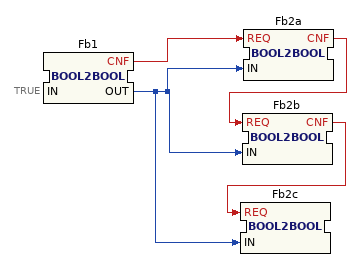
      [picture p24: application _03_DataConnections.Ex2b]
      FBS
        Fb1 : BOOL2BOOL(IN := TRUE);
        Fb2a : BOOL2BOOL;
        Fb2b : BOOL2BOOL;
        Fb2c : BOOL2BOOL;
      END_FBS
      EVENT_CONNECTIONS
        Fb1.CNF TO Fb2a.REQ;
        Fb2a.CNF TO Fb2b.REQ;
        Fb2b.CNF TO Fb2c.REQ;
      END_CONNECTIONS
      DATA_CONNECTIONS
        Fb1.OUT TO Fb2a.IN;
        Fb1.OUT TO Fb2b.IN;
        Fb1.OUT TO Fb2c.IN;
      END_CONNECTIONS
    END_SUBAPPLICATION
    SUBAPPLICATION Ex4b (* type casts (explicit, downcast) &#10;- trigger Fb1.REQ &#10;- expect Fb3.CUO and CV:=1 and Q:=TRUE *)
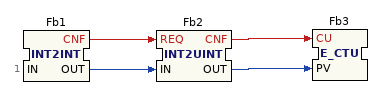
      FBS
        Fb1 : INT2INT(IN := 1);
        Fb3 : E_CTU;
        Fb2 : INT2UINT;
      END_FBS
      EVENT_CONNECTIONS
        Fb1.CNF TO Fb2.REQ;
        Fb2.CNF TO Fb3.CU;
      END_CONNECTIONS
      DATA_CONNECTIONS
        Fb1.OUT TO Fb2.IN;
        Fb2.OUT TO Fb3.PV;
      END_CONNECTIONS
    END_SUBAPPLICATION
    SUBAPPLICATION Ex5a (* type casts (implicit, upcast from UINT to LREAL) &#10;- trigger Fb1.CU  &#10;- expect Fb2.CNF and Fb2.OUT:=INT#6 *)
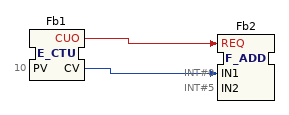
      FBS
        Fb1 : E_CTU(PV := 10);
        Fb2 : F_ADD(IN1 := INT#0, IN2 := INT#5);
      END_FBS
      EVENT_CONNECTIONS
        Fb1.CUO TO Fb2.REQ;
      END_CONNECTIONS
      DATA_CONNECTIONS
        Fb1.CV TO Fb2.IN1;
      END_CONNECTIONS
    END_SUBAPPLICATION
    SUBAPPLICATION Ex5b (* type casts (implicit, upcast from UINT to ANY_MAG) &#10;- trigger Fb1.CU &#10;- expect Fb2.CNF and Fb2.OUT:=REAL#1.0 *)
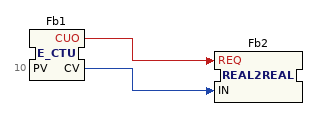
      FBS
        Fb1 : E_CTU(PV := 10);
        Fb2 : REAL2REAL;
      END_FBS
      EVENT_CONNECTIONS
        Fb1.CUO TO Fb2.REQ;
      END_CONNECTIONS
      DATA_CONNECTIONS
        Fb1.CV TO Fb2.IN;
      END_CONNECTIONS
    END_SUBAPPLICATION
  END_APPLICATION
  APPLICATION _07_Subapplications
    (* Group __Group01: connection to the interface *)
  END_APPLICATION
  APPLICATION _06_CompositeFBs
    (* Group __Group01: WITH bei composite FBs *)
  END_APPLICATION
  APPLICATION _02_Parameters
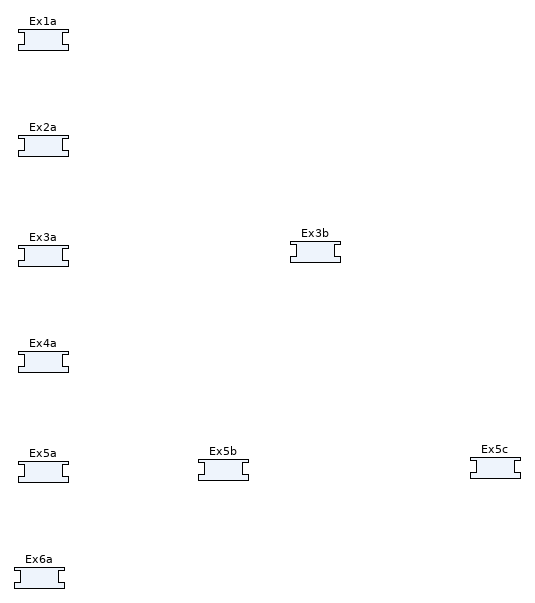
    (* Group Info_Parameters: The subapps in this App serve as test cases for various versions of parameters: &#10;- simple boolean parameters (including counter-examples) &#10;- initial value taken from type when no parameter is present &#10;- parameters with prefixes &#10;- upcasts in parameters *)
    SUBAPPLICATION Ex2a (* Parameters &#10; &#10;- Trigger EI  &#10;- Expect nothing *)
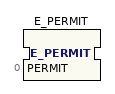
      FBS
        E_PERMIT : E_PERMIT(PERMIT := 0);
      END_FBS
    END_SUBAPPLICATION
    SUBAPPLICATION Ex1a (* Parameters overriding initial value of data type &#10; &#10;- Trigger E_PERMIT.EI  &#10;- Expect E_PERMIT.EO *)
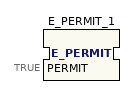
      FBS
        E_PERMIT_1 : E_PERMIT(PERMIT := TRUE);
      END_FBS
    END_SUBAPPLICATION
    SUBAPPLICATION Ex3a (* Initial Value (from type) &#10; &#10;- Trigger EI  &#10;- Expect EO *)
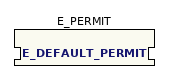
      FBS
        E_PERMIT : E_DEFAULT_PERMIT;
      END_FBS
    END_SUBAPPLICATION
    SUBAPPLICATION Ex4a (* Override initial value (from type) with parameter &#10; &#10;- Trigger EI  &#10;- Expect nothing *)
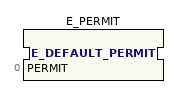
      FBS
        E_PERMIT : E_DEFAULT_PERMIT(PERMIT := 0);
      END_FBS
    END_SUBAPPLICATION
    SUBAPPLICATION Ex6a (* Any type: required casts  &#10; &#10;- Trigger REQ &#10;- Expect CNF and OUT:=13 *)
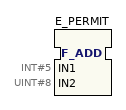
      FBS
        E_PERMIT : F_ADD(IN1 := INT#5, IN2 := UINT#8);
      END_FBS
    END_SUBAPPLICATION
    SUBAPPLICATION Ex5a (* integer parameter &#10; &#10;- Trigger REQ &#10;- Expect CNF, OUT:=5 *)
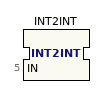
      FBS
        INT2INT : INT2INT(IN := 5);
      END_FBS
    END_SUBAPPLICATION
    SUBAPPLICATION Ex5b (* integer parameter with prefix &#10; &#10;- Trigger REQ &#10;- Expect CNF, OUT:=5 *)
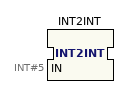
      FBS
        INT2INT : INT2INT(IN := INT#5);
      END_FBS
    END_SUBAPPLICATION
    SUBAPPLICATION Ex5c (* integer parameter with prefix (upcast) &#10; &#10;- Trigger REQ &#10;- Expect CNF, OUT:=5 *)
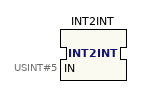
      FBS
        INT2INT : INT2INT(IN := USINT#5);
      END_FBS
    END_SUBAPPLICATION
    SUBAPPLICATION Ex3b (* Initial Value (from type)  &#10;  &#10;- Trigger EI   &#10;- Expect nothing *)
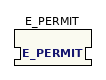
      FBS
        E_PERMIT : E_PERMIT;
      END_FBS
    END_SUBAPPLICATION
  END_APPLICATION
  APPLICATION _04_DataWith
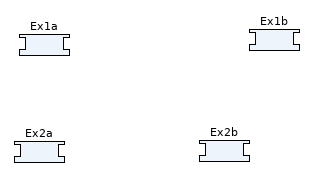
    (* Group Info_DataConnections: The subapps in this App serve as test cases for various versions of WITH-constructs (on updating data values to the outputs). &#10;- WITH at the inputs &#10;- WITH at the outputs *)
    SUBAPPLICATION Ex1a (* no WITH at the output variables, do not update &#10;trigger REQ, expect CNF and  &#10;DO1.OUT:=TRUE  &#10;DO2.OUT:=-10  &#10;DO3.OUT:=15  &#10;DO4.OUT:=2.0 (data values from type) *)
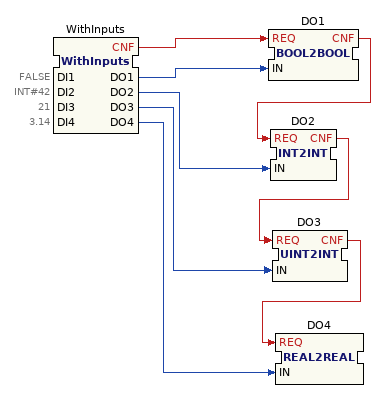
      FBS
        WithInputs : WithInputs(DI1 := FALSE, DI2 := INT#42, DI3 := 21, DI4 := 3.14);
        DO1 : BOOL2BOOL;
        DO2 : INT2INT;
        DO3 : UINT2INT;
        DO4 : REAL2REAL;
      END_FBS
      EVENT_CONNECTIONS
        WithInputs.CNF TO DO1.REQ;
        DO1.CNF TO DO2.REQ;
        DO2.CNF TO DO3.REQ;
        DO3.CNF TO DO4.REQ;
      END_CONNECTIONS
      DATA_CONNECTIONS
        WithInputs.DO1 TO DO1.IN;
        WithInputs.DO2 TO DO2.IN;
        WithInputs.DO3 TO DO3.IN;
        WithInputs.DO4 TO DO4.IN;
      END_CONNECTIONS
    END_SUBAPPLICATION
    SUBAPPLICATION Ex1b (* WITH at the output values, update &#10;trigger UPDATE, expect CNF and   &#10;DO1.OUT:=FALSE   &#10;DO2.OUT:=42   &#10;DO3.OUT:=21   &#10;DO4.OUT:=3.14 (data values from instance) *)
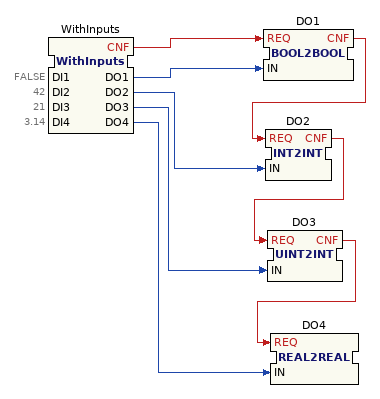
      FBS
        WithInputs : WithInputs(DI1 := FALSE, DI2 := 42, DI3 := 21, DI4 := 3.14);
        DO1 : BOOL2BOOL;
        DO2 : INT2INT;
        DO3 : UINT2INT;
        DO4 : REAL2REAL;
      END_FBS
      EVENT_CONNECTIONS
        WithInputs.CNF TO DO1.REQ;
        DO1.CNF TO DO2.REQ;
        DO2.CNF TO DO3.REQ;
        DO3.CNF TO DO4.REQ;
      END_CONNECTIONS
      DATA_CONNECTIONS
        WithInputs.DO1 TO DO1.IN;
        WithInputs.DO2 TO DO2.IN;
        WithInputs.DO3 TO DO3.IN;
        WithInputs.DO4 TO DO4.IN;
      END_CONNECTIONS
    END_SUBAPPLICATION
    SUBAPPLICATION Ex2a (* trigger REQ, expect CNF and  &#10;DO1.OUT:=TRUE  &#10;DO2.OUT:=-42  &#10;DO3.OUT:=21  &#10;DO4.OUT:=0.0 (data values from type) *)
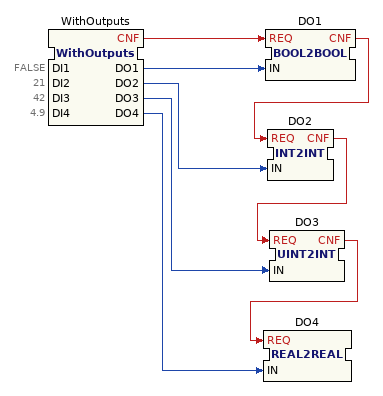
      FBS
        DO1 : BOOL2BOOL;
        DO2 : INT2INT;
        DO3 : UINT2INT;
        DO4 : REAL2REAL;
        WithOutputs : WithOutputs(DI1 := FALSE, DI2 := 21, DI3 := 42, DI4 := 4.9);
      END_FBS
      EVENT_CONNECTIONS
        DO1.CNF TO DO2.REQ;
        DO2.CNF TO DO3.REQ;
        DO3.CNF TO DO4.REQ;
        WithOutputs.CNF TO DO1.REQ;
      END_CONNECTIONS
      DATA_CONNECTIONS
        WithOutputs.DO1 TO DO1.IN;
        WithOutputs.DO2 TO DO2.IN;
        WithOutputs.DO3 TO DO3.IN;
        WithOutputs.DO4 TO DO4.IN;
      END_CONNECTIONS
    END_SUBAPPLICATION
    SUBAPPLICATION Ex2b (* trigger UPDATE, expect CNF and &#10;DO1.OUT:=FALSE &#10;DO2.OUT:=21 &#10;DO3.OUT:=42 &#10;DO4.OUT:=4.9 (data values from parameters) *)
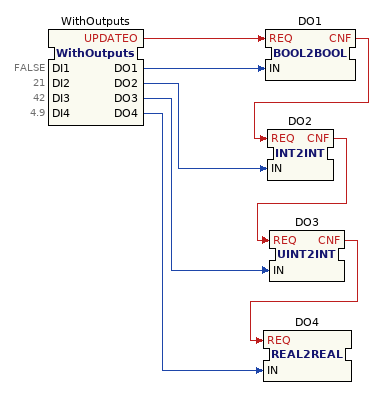
      FBS
        DO1 : BOOL2BOOL;
        DO2 : INT2INT;
        DO3 : UINT2INT;
        DO4 : REAL2REAL;
        WithOutputs : WithOutputs(DI1 := FALSE, DI2 := 21, DI3 := 42, DI4 := 4.9);
      END_FBS
      EVENT_CONNECTIONS
        DO1.CNF TO DO2.REQ;
        DO2.CNF TO DO3.REQ;
        DO3.CNF TO DO4.REQ;
        WithOutputs.UPDATEO TO DO1.REQ;
      END_CONNECTIONS
      DATA_CONNECTIONS
        WithOutputs.DO1 TO DO1.IN;
        WithOutputs.DO2 TO DO2.IN;
        WithOutputs.DO3 TO DO3.IN;
        WithOutputs.DO4 TO DO4.IN;
      END_CONNECTIONS
    END_SUBAPPLICATION
  END_APPLICATION
  APPLICATION _05_Adapter
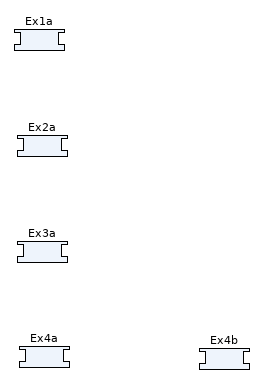
    (* Group Info_Adapter: The subapps in this App serve as test cases for various versions of WITH-constructs (on updating data values to the outputs). &#10;- WITH at the inputs &#10;- WITH at the outputs *)
    SUBAPPLICATION Ex1a (* Adapter with just events &#10;- trigger Fb1.REQ  &#10;- expect Fb1.CNF and Fb1.RSP *)
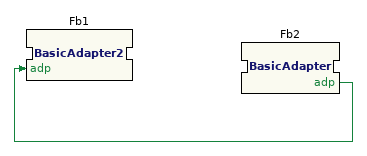
      FBS
        Fb1 : BasicAdapter2;
        Fb2 : BasicAdapter;
      END_FBS
      ADAPTER_CONNECTIONS
        Fb2.adp TO Fb1.adp;
      END_CONNECTIONS
    END_SUBAPPLICATION
    SUBAPPLICATION Ex2a (* Adapter with an event and data  &#10;- trigger Fb1.REQ   &#10;- expect Fb2.CNF with Fb2.DO1 := 5, Fb2.DO2 := TRUE *)
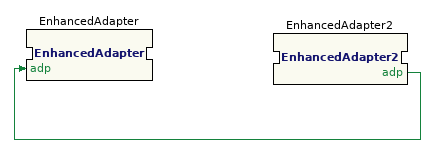
      FBS
        EnhancedAdapter : EnhancedAdapter;
        EnhancedAdapter2 : EnhancedAdapter2;
      END_FBS
      ADAPTER_CONNECTIONS
        EnhancedAdapter2.adp TO EnhancedAdapter.adp;
      END_CONNECTIONS
    END_SUBAPPLICATION
    SUBAPPLICATION Ex3a (* Adapter with a WITH (do not update all data)  &#10;- trigger Fb1.REQ   &#10;- expect Fb2.CNF with Fb2.DO1 := 5, Fb2.DO2 := FALSE *)
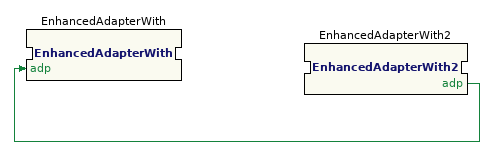
      FBS
        EnhancedAdapterWith2 : EnhancedAdapterWith2;
        EnhancedAdapterWith : EnhancedAdapterWith;
      END_FBS
      ADAPTER_CONNECTIONS
        EnhancedAdapterWith2.adp TO EnhancedAdapterWith.adp;
      END_CONNECTIONS
    END_SUBAPPLICATION
    SUBAPPLICATION Ex4a (* analyze default values of adapter &#10;trigger REQ &#10;outputs show the 4 default values of the adapter *)
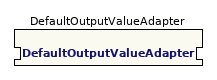
      FBS
        DefaultOutputValueAdapter : DefaultOutputValueAdapter;
      END_FBS
    END_SUBAPPLICATION
    SUBAPPLICATION Ex4b (* analyze default values of adapter &#10;trigger REQ &#10;outputs show the 4 default values of the adapter *)
